Universal Robots URScript: ManyMoves.script

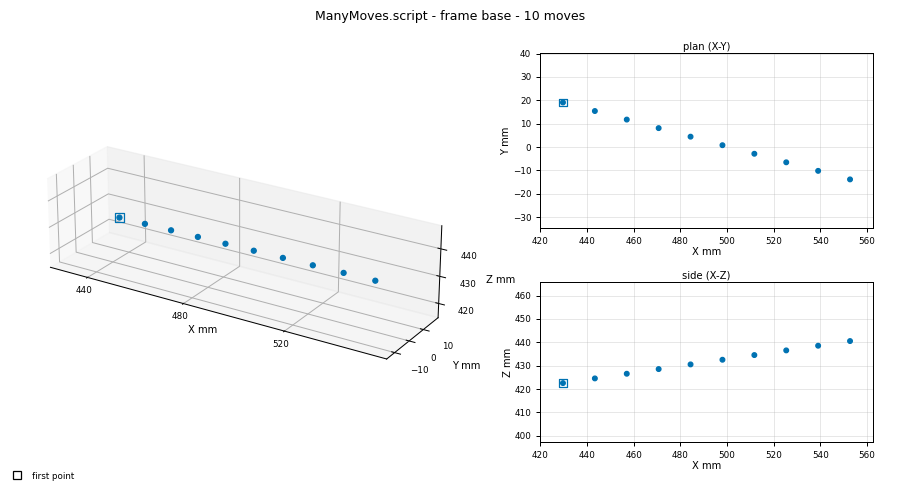
[picture p0: tool path of ManyMoves.script in frame base, 10 of 40 moves have a stored position in this frame; points joined in program order, loops and branches not executed]
def ManyMoves():
  # Global parameters:
  global speed_ms    = 0.250
  global speed_rads  = 0.750
  global accel_mss   = 1.200
  global accel_radss = 1.200
  global blend_radius_m = 0.001
  global ref_frame = p[0,0,0,0,0,0]

  #
  # TO REMOVE HEADER:
  # Go to "Program" -> "Post-Processor Editor"
  # Select "Universal Robots"
  # Set "INCLUDE_HEADER" to "False"
  #
  #--------------------------
  # Add any default subprograms here
  # For example, to drive a gripper as a program call:
  # def Gripper_Open():
  #   ...
  # end
  #
  # Example to drive a spray gun:
  def SprayOn(value):
    # use the value as an output:
    DO_SPRAY = 5
    if value == 0:
      set_standard_digital_out(DO_SPRAY, False)
    else:
      set_standard_digital_out(DO_SPRAY, True)
    end
  end

  # Example to drive an extruder:
  def Extruder(value):
    # use the value as an output:
    if value < 0:
      # stop extruder
    else:
      # start extruder
    end
  end

  # Example to move an external axis
  def MoveAxis(value):
    # use the value as an output:
    DO_AXIS_1 = 1
    DI_AXIS_1 = 1
    if value <= 0:
      set_standard_digital_out(DO_AXIS_1, False)

      # Wait for digital input to change state
      #while (get_standard_digital_in(DI_AXIS_1) != False):
      #  sync()
      #end
    else:
      set_standard_digital_out(DO_AXIS_1, True)

      # Wait for digital input to change state
      #while (get_standard_digital_in(DI_AXIS_1) != True):
      #  sync()
      #end
    end
  end
  #--------------------------


  # Main program:
  # Program generated by RoboDK v6.0.7 for UR10 on XX/XX/XXXX 18:00:00
  # Using nominal kinematics.
  ref_frame = p[1.234570, -0.098765, 0.050500, 0.000000, 0.000000, 0.523599]
  set_tcp(p[0.010000, 0.020000, 0.150000, 0.000000, 0.000000, 0.000000])
  speed_ms    = 0.500
  movej([0.000000, -0.174533, 0.349066, 0.000000, 0.523599, 0.000000],accel_radss,speed_rads,t=0,r=0)
  movel(pose_trans(ref_frame,p[-0.638084, 0.504480, 0.372034, 0.731956, 2.185937, -0.570291]),accel_mss,speed_ms,t=0,r=0.001)
  movej([0.349066, -0.174533, 0.349066, 0.000000, 0.523599, 0.000000],accel_radss,speed_rads,t=0,r=0)
  movel([0.000000, -0.174533, 0.349066, 0.000000, 0.523599, 0.000000],accel_mss,speed_ms,t=0,r=0)
  movej([0.000000, -0.174533, 0.349066, 0.000000, 0.523599, 0.000000],accel_radss,speed_rads,t=0,r=0)
  movel(pose_trans(ref_frame,p[-0.628084, 0.494480, 0.374034, 0.731956, 2.185937, -0.570291]),accel_mss,speed_ms,t=0,r=0.001)
  movej([0.349066, -0.174533, 0.349066, 0.000000, 0.523599, 0.000000],accel_radss,speed_rads,t=0,r=0)
  movel([0.000000, -0.174533, 0.349066, 0.000000, 0.523599, 0.000000],accel_mss,speed_ms,t=0,r=0)
  movej([0.000000, -0.174533, 0.349066, 0.000000, 0.523599, 0.000000],accel_radss,speed_rads,t=0,r=0)
  movel(pose_trans(ref_frame,p[-0.618084, 0.484480, 0.376034, 0.731956, 2.185937, -0.570291]),accel_mss,speed_ms,t=0,r=0.001)
  movej([0.349066, -0.174533, 0.349066, 0.000000, 0.523599, 0.000000],accel_radss,speed_rads,t=0,r=0)
  movel([0.000000, -0.174533, 0.349066, 0.000000, 0.523599, 0.000000],accel_mss,speed_ms,t=0,r=0)
  movej([0.000000, -0.174533, 0.349066, 0.000000, 0.523599, 0.000000],accel_radss,speed_rads,t=0,r=0)
  movel(pose_trans(ref_frame,p[-0.608084, 0.474480, 0.378034, 0.731956, 2.185937, -0.570291]),accel_mss,speed_ms,t=0,r=0.001)
  movej([0.349066, -0.174533, 0.349066, 0.000000, 0.523599, 0.000000],accel_radss,speed_rads,t=0,r=0)
  movel([0.000000, -0.174533, 0.349066, 0.000000, 0.523599, 0.000000],accel_mss,speed_ms,t=0,r=0)
  movej([0.000000, -0.174533, 0.349066, 0.000000, 0.523599, 0.000000],accel_radss,speed_rads,t=0,r=0)
  movel(pose_trans(ref_frame,p[-0.598084, 0.464480, 0.380034, 0.731956, 2.185937, -0.570291]),accel_mss,speed_ms,t=0,r=0.001)
  movej([0.349066, -0.174533, 0.349066, 0.000000, 0.523599, 0.000000],accel_radss,speed_rads,t=0,r=0)
  movel([0.000000, -0.174533, 0.349066, 0.000000, 0.523599, 0.000000],accel_mss,speed_ms,t=0,r=0)
  movej([0.000000, -0.174533, 0.349066, 0.000000, 0.523599, 0.000000],accel_radss,speed_rads,t=0,r=0)
  movel(pose_trans(ref_frame,p[-0.588084, 0.454480, 0.382034, 0.731956, 2.185937, -0.570291]),accel_mss,speed_ms,t=0,r=0.001)
  movej([0.349066, -0.174533, 0.349066, 0.000000, 0.523599, 0.000000],accel_radss,speed_rads,t=0,r=0)
  movel([0.000000, -0.174533, 0.349066, 0.000000, 0.523599, 0.000000],accel_mss,speed_ms,t=0,r=0)
  movej([0.000000, -0.174533, 0.349066, 0.000000, 0.523599, 0.000000],accel_radss,speed_rads,t=0,r=0)
  movel(pose_trans(ref_frame,p[-0.578084, 0.444480, 0.384034, 0.731956, 2.185937, -0.570291]),accel_mss,speed_ms,t=0,r=0.001)
  movej([0.349066, -0.174533, 0.349066, 0.000000, 0.523599, 0.000000],accel_radss,speed_rads,t=0,r=0)
  movel([0.000000, -0.174533, 0.349066, 0.000000, 0.523599, 0.000000],accel_mss,speed_ms,t=0,r=0)
  movej([0.000000, -0.174533, 0.349066, 0.000000, 0.523599, 0.000000],accel_radss,speed_rads,t=0,r=0)
  movel(pose_trans(ref_frame,p[-0.568084, 0.434480, 0.386034, 0.731956, 2.185937, -0.570291]),accel_mss,speed_ms,t=0,r=0.001)
  movej([0.349066, -0.174533, 0.349066, 0.000000, 0.523599, 0.000000],accel_radss,speed_rads,t=0,r=0)
  movel([0.000000, -0.174533, 0.349066, 0.000000, 0.523599, 0.000000],accel_mss,speed_ms,t=0,r=0)
  movej([0.000000, -0.174533, 0.349066, 0.000000, 0.523599, 0.000000],accel_radss,speed_rads,t=0,r=0)
  movel(pose_trans(ref_frame,p[-0.558084, 0.424480, 0.388034, 0.731956, 2.185937, -0.570291]),accel_mss,speed_ms,t=0,r=0.001)
  movej([0.349066, -0.174533, 0.349066, 0.000000, 0.523599, 0.000000],accel_radss,speed_rads,t=0,r=0)
  movel([0.000000, -0.174533, 0.349066, 0.000000, 0.523599, 0.000000],accel_mss,speed_ms,t=0,r=0)
  movej([0.000000, -0.174533, 0.349066, 0.000000, 0.523599, 0.000000],accel_radss,speed_rads,t=0,r=0)
  movel(pose_trans(ref_frame,p[-0.548084, 0.414480, 0.390034, 0.731956, 2.185937, -0.570291]),accel_mss,speed_ms,t=0,r=0.001)
  movej([0.349066, -0.174533, 0.349066, 0.000000, 0.523599, 0.000000],accel_radss,speed_rads,t=0,r=0)
  movel([0.000000, -0.174533, 0.349066, 0.000000, 0.523599, 0.000000],accel_mss,speed_ms,t=0,r=0)
  # End of main program
end

ManyMoves()
